// TIA Portal project "Robotic_arm" (V19)

(* hardware
DEVICE "S7-1500/ET200MP station_1"  S7-1500 station
   slot 0: "Rail_0"  Rack  6ES7 590-1***0-0AA0
   slot 1: "PLC_2"  CPU 1511-1 PN  6ES7 511-1AK00-0AB0  V1.8
      slot 3: "CPU display_1"  6ES7591-1AA00-0AA0
      slot 32768: "PROFINET interface_1"  X1
         slot 32769: "Port_1"  X1 P1
         slot 32770: "Port_2"  X1 P2
*)

// ===== PLC "PLC_2"  CPU 1511-1 PN =====

VAR_GLOBAL   // PLC tag table "Cell_IO_list"
   "Cmd_Band_Run" AT %Q0.0 : Bool;
   "Cmd_Gripper_Close" AT %Q0.1 : Bool;
   "Cmd_LoadNew" AT %Q0.2 : Bool;
   "Cmd_Picked" AT %Q0.3 : Bool;
   "Cmd_A1_Pos" AT %QD4 : Real;
   "Cmd_A2_Pos" AT %QD8 : Real;
   "Cmd_A3_Pos" AT %QD12 : Real;
   "Cmd_A4_Pos" AT %QD16 : Real;
   "St_ProductAtPick" AT %I1.0 : Bool;
   "St_Gripper_HasPart" AT %I1.1 : Bool;
   "St_A1_Pos" AT %ID4 : Real;
   "St_A2_Pos" AT %ID8 : Real;
   "St_A3_Pos" AT %ID12 : Real;
   "St_A4_Pos" AT %ID16 : Real;
   "Cmd_Start" AT %M0.0 : Bool;
   "Cmd_Stop" AT %M0.1 : Bool;
   "Cmd_Reset" AT %M0.2 : Bool;
   "Cmd_Auto" AT %M0.3 : Bool;
   "SafeToRun" AT %M0.4 : Bool;
   "Sts_Ready" AT %M10.0 : Bool;
   "Sts_Busy" AT %M10.1 : Bool;
   "Sts_Done" AT %M10.2 : Bool;
   "Sts_Fault" AT %M10.3 : Bool;
   "Sts_State" AT %MW12 : Int;
   "Sts_CycleCount" AT %MW14 : Int;
   "Sts_Hold" AT %M10.4 : Bool;
END_VAR

DATA_BLOCK "DB_RobotPoses"   // DB1
{ S7_Optimized_Access := 'TRUE' }
VERSION : 0.3
   VAR
      HOME_A1 : Real;
      HOME_A2 : Real;
      HOME_A3 : Real;
      HOME_A4 : Real;
      PICK_APP_A1 : Real;
      PICK_APP_A2 : Real := -31.0;
      PICK_APP_A3 : Real := -28.6;
      PICK_APP_A4 : Real := 59.6;
      PICK_A1 : Real;
      PICK_A2 : Real := -50.8;
      PICK_A3 : Real := -24.4;
      PICK_A4 : Real := 75.2;
      PLACE_APP_A1 : Real := 90.0;
      PLACE_APP_A2 : Real := -5.4;
      PLACE_APP_A3 : Real := -51.3;
      PLACE_APP_A4 : Real := 56.7;
      PLACE_A1 : Real := 90.0;
      PLACE_A2 : Real := -42.1;
      PLACE_A3 : Real := -48.1;
      PLACE_A4 : Real := 90.2;
   END_VAR
BEGIN
END_DATA_BLOCK

DATA_BLOCK "iCell"   // DB6
{ S7_Optimized_Access := 'TRUE' }
VERSION : 0.3
// stored: InstanceOfName FB_CellController
"FB_CellController"
BEGIN
END_DATA_BLOCK

FUNCTION_BLOCK "FB_RobotMove"   // FB1, SCL
{ S7_Optimized_Access := 'TRUE' }
VERSION : 0.5
// ----------------------------------------------------------------------------
//  FB_RobotMove : command one joint pose, report Done from NX actual positions
//    - writes the 4 joint set-points to NX (Cmd*)
//    - Done when every joint is within Tol of its target AND a minimum settle
//      time has elapsed.
// 
//    FIX 1: the move re-arms on a rising edge of Execute OR whenever the caller's
//    Step number changes.  The caller passes its own CASE state as Step, so every
//    state transition starts a genuinely new move even when Execute stays TRUE and
//    even when two consecutive states share the same target pose.
//  ----------------------------------------------------------------------------
   VAR_INPUT
      Execute : Bool;
      "Step" : Int;   // caller's state number (FIX 1)
      T1 : Real;   // target joint angles
      T2 : Real;
      T3 : Real;
      T4 : Real;
      Act1 : Real;   // actual angles from NX
      Act2 : Real;
      Act3 : Real;
      Act4 : Real;
      Tol : Real;   // tolerance [deg]
   END_VAR
   VAR_OUTPUT
      Cmd1 : Real := 0.0;   // set-points to NX
      Cmd2 : Real := 0.0;
      Cmd3 : Real := 0.0;
      Cmd4 : Real := 0.0;
      Done : Bool := FALSE;
      Busy : Bool := FALSE;
   END_VAR
   VAR
      prevExec : Bool;
      iBusy : Bool := FALSE;   // FIX 9: internal, so no output is read
      prevStep : Int := -1;
      SettleT : TON_TIME;
   END_VAR
   VAR_TEMP
      inpos : Bool;
      startMove : Bool;
   END_VAR
BEGIN

   // ---- start a new move: rising Execute, or the caller moved to a new step ----
   #startMove := #Execute AND ((NOT #prevExec) OR (#Step <> #prevStep));       // FIX 1

   IF #startMove THEN
       #iBusy := TRUE;
       #Done := FALSE;
   END_IF;

   #prevExec := #Execute;
   #prevStep := #Step;

   // drive set-points only while this move is selected
   IF #Execute THEN
       #Cmd1 := #T1;
       #Cmd2 := #T2;
       #Cmd3 := #T3;
       #Cmd4 := #T4;
   END_IF;

   // in-position test on the NX feedback
   #inpos := (ABS(#Act1 - #T1) <= #Tol) AND
   (ABS(#Act2 - #T2) <= #Tol) AND
   (ABS(#Act3 - #T3) <= #Tol) AND
   (ABS(#Act4 - #T4) <= #Tol);

   // minimum settle / move time.
   // FIX 2: held at IN := FALSE for the re-arm scan, which resets the TON, so the
   //        settle time is honoured for EVERY move and not just the first one.
   #SettleT(IN := #iBusy AND NOT #startMove,
            PT := T#200ms);

   IF #iBusy AND #inpos AND #SettleT.Q THEN
       #Done := TRUE;
       #iBusy := FALSE;
   END_IF;

   // deselecting the move clears it
   IF NOT #Execute THEN
       #Done := FALSE;
       #iBusy := FALSE;
       #prevStep := -1;
   END_IF;

   #Busy := #iBusy;
END_FUNCTION_BLOCK

FUNCTION_BLOCK "FB_Geven"   // FB2, SCL
{ S7_Optimized_Access := 'TRUE' }
VERSION : 0.5
// ----------------------------------------------------------------------------
//  FB_Geven  (GIVE) : run the conveyor until the product reaches the pick
//                     light barrier, then stop the belt. Fault on arrival
//                     time-out (product never arrives).
//    INTERLOCK: the belt only ever runs from inside this module.
//  ----------------------------------------------------------------------------
   VAR_INPUT
      Run : Bool;   // enabled by CellController (active AND not held)
      SafeToRun : Bool;
      St_ProductAtPick : Bool;
   END_VAR
   VAR_OUTPUT
      Cmd_Band_Run : Bool := FALSE;
      Done : Bool := FALSE;
      Fault : Bool := FALSE;
   END_VAR
   VAR
      ArriveTO : TON_TIME;
      iFault : Bool := FALSE;   // FIX 9
      iBand : Bool := FALSE;   // FIX 9
      Cleared : Bool := FALSE;   // FIX 10: barrier seen clear since this module started
   END_VAR
BEGIN

   IF #Run AND #SafeToRun AND NOT #iFault THEN
       IF NOT #Cleared THEN
           // FIX 10: on entry the light barrier may STILL be showing the previous
           //         product (the status signal is one communication step old).
           //         Feed, but do not accept an arrival until the barrier has been
           //         seen clear at least once, so a stale TRUE cannot be mistaken
           //         for the next product arriving.
           #iBand := TRUE;
           #Done := FALSE;
           IF NOT #St_ProductAtPick THEN
               #Cleared := TRUE;
           END_IF;
       ELSIF #St_ProductAtPick THEN
           #iBand := FALSE;     // product detected -> stop belt (pick interlock)
           #Done := TRUE;
       ELSE
           #iBand := TRUE;      // keep feeding
           #Done := FALSE;
       END_IF;
   ELSE
       #iBand := FALSE;
   END_IF;

   // arrival time-out -> representative process error.
   // Called every scan; IN follows the belt command, so it resets by itself when
   // the belt stops or when the module is deselected.
   #ArriveTO(IN := #iBand,
             PT := T#15s);
   IF #ArriveTO.Q THEN
       #iFault := TRUE;
       #iBand := FALSE;
   END_IF;

   IF NOT #Run THEN                  // reset when CellController deselects the module
       #Done := FALSE;
       #iFault := FALSE;
       #Cleared := FALSE;             // FIX 10: re-arm for the next cycle
   END_IF;

   #Cmd_Band_Run := #iBand;
   #Fault := #iFault;
END_FUNCTION_BLOCK

FUNCTION_BLOCK "FB_Verwerken"   // FB3, SCL
{ S7_Optimized_Access := 'TRUE' }
VERSION : 0.3
// RobotCell v0.3 PATCH - only the two blocks that change (FIX 6).
//  FB_RobotMove, FB_Geven, FB_Wegzetten and DB_RobotPoses stay as they are in TIA.
//  ----------------------------------------------------------------------------
//  FB_Verwerken  (PROCESS) : robot picks the product.
//    PICK_APP -> PICK -> close gripper (wait HasPart + 0.5 s) -> lift to PICK_APP
//    -> check the presence sensor is clear (FIX 6).  Missed pick -> retry (max 2).
//    Fault on grip time-out (no part after closing) or on the third missed pick.
//  ----------------------------------------------------------------------------
   VAR_INPUT
      Run : Bool;
      SafeToRun : Bool;
      Act1 : Real;
      Act2 : Real;
      Act3 : Real;
      Act4 : Real;
      St_Gripper_HasPart : Bool;
      St_ProductAtPick : Bool;   // FIX 6: presence sensor at the pick point
   END_VAR
   VAR_OUTPUT
      Cmd1 : Real;
      Cmd2 : Real;
      Cmd3 : Real;
      Cmd4 : Real;
      Cmd_Gripper_Close : Bool;
      Done : Bool;
      Fault : Bool;
      Retries : Int;   // FIX 6: missed picks in this cycle
   END_VAR
   VAR
      State : Int := 0;
      Move : "FB_RobotMove";
      GripTO : TON_TIME;
      GripSettle : TON_TIME;   // FIX 6: jaws settle before lifting
      CheckT : TON_TIME;   // FIX 6: sensor settle after the lift
   END_VAR
BEGIN
   // =====================================================================
   // FB_Verwerken  v0.3  -  CODE ONLY (paste into the code area, replace all)
   //
   // Before pasting, add these 4 lines to the INTERFACE table at the top:
   //   Input   St_ProductAtPick   Bool
   //   Output  Retries            Int
   //   Static  GripSettle         TON_TIME
   //   Static  CheckT             TON_TIME
   // (Run, SafeToRun, Act1..Act4, St_Gripper_HasPart, Cmd1..Cmd4,
   //  Cmd_Gripper_Close, Done, Fault, State, Move, GripTO stay as they are.)
   // =====================================================================

   // FIX 3: the grip time-out is called ONCE PER SCAN, outside the CASE, with an
   //        explicit enable.  It therefore sees IN = FALSE whenever the module is
   //        idle or in another step, which resets it between cycles.  In v0.1 it
   //        was only called from inside CASE 20 with IN := TRUE and kept its
   //        elapsed time, so cycle 2 faulted immediately on entry.
   #GripTO(IN := #Run AND #SafeToRun AND NOT #Fault AND (#State = 20),
           PT := T#3s);
   #GripSettle(IN := #Run AND #SafeToRun AND (#State = 20) AND #St_Gripper_HasPart,
               PT := T#500ms);
   #CheckT(IN := #Run AND #SafeToRun AND (#State = 40),
           PT := T#300ms);

   IF NOT #Run THEN
       #State := 0;
       #Done := FALSE;
       #Fault := FALSE;
       #Retries := 0;
       #Cmd_Gripper_Close := FALSE;
       #Move(Execute := FALSE,
             Step := -1,
             Tol := 1.0,
             Act1 := #Act1,
             Act2 := #Act2,
             Act3 := #Act3,
             Act4 := #Act4);
   ELSIF #SafeToRun AND NOT #Fault THEN
       CASE #State OF
           0:  // move to PICK approach
               #Move(Execute := TRUE,
                     Step := 0,
                     Tol := 1.0,
                     T1 := "DB_RobotPoses".PICK_APP_A1,
                     T2 := "DB_RobotPoses".PICK_APP_A2,
                     T3 := "DB_RobotPoses".PICK_APP_A3,
                     T4 := "DB_RobotPoses".PICK_APP_A4,
                     Act1 := #Act1,
                     Act2 := #Act2,
                     Act3 := #Act3,
                     Act4 := #Act4);
               IF #Move.Done THEN
                   #State := 10;
               END_IF;

           10: // descend to PICK
               #Move(Execute := TRUE,
                     Step := 10,
                     Tol := 1.0,
                     T1 := "DB_RobotPoses".PICK_A1,
                     T2 := "DB_RobotPoses".PICK_A2,
                     T3 := "DB_RobotPoses".PICK_A3,
                     T4 := "DB_RobotPoses".PICK_A4,
                     Act1 := #Act1,
                     Act2 := #Act2,
                     Act3 := #Act3,
                     Act4 := #Act4);
               IF #Move.Done THEN
                   #State := 20;
               END_IF;

           20: // close gripper, wait for part, let the jaws settle (FIX 6)
               #Cmd_Gripper_Close := TRUE;
               IF #GripSettle.Q THEN
                   #State := 30;
               ELSIF #GripTO.Q THEN
                   #Fault := TRUE;            // grip time-out -> error
               END_IF;

           30: // lift back to PICK approach (with part)
               #Move(Execute := TRUE,
                     Step := 30,
                     Tol := 1.0,
                     T1 := "DB_RobotPoses".PICK_APP_A1,
                     T2 := "DB_RobotPoses".PICK_APP_A2,
                     T3 := "DB_RobotPoses".PICK_APP_A3,
                     T4 := "DB_RobotPoses".PICK_APP_A4,
                     Act1 := #Act1,
                     Act2 := #Act2,
                     Act3 := #Act3,
                     Act4 := #Act4);
               IF #Move.Done THEN
                   #State := 40;
               END_IF;

           40: // FIX 6: verify the pick with the presence sensor
               IF #CheckT.Q THEN
                   IF NOT #St_ProductAtPick THEN
                       #State := 100;          // block left the belt -> picked
                   ELSIF #Retries < 2 THEN
                       #Retries := #Retries + 1; // block still there -> missed pick
                       #Cmd_Gripper_Close := FALSE;
                       #State := 50;
                   ELSE
                       #Fault := TRUE;         // third miss -> process error
                   END_IF;
               END_IF;

           50: // FIX 6: retry - open above the block, then descend again
               #Cmd_Gripper_Close := FALSE;
               IF NOT #St_Gripper_HasPart THEN
                   #State := 10;
               END_IF;

           100: // done
               #Done := TRUE;
       END_CASE;
   END_IF;

   // hand the move set-points to the block outputs (read by FB_CellController in step 20)
   #Cmd1 := #Move.Cmd1;
   #Cmd2 := #Move.Cmd2;
   #Cmd3 := #Move.Cmd3;
   #Cmd4 := #Move.Cmd4;
END_FUNCTION_BLOCK

FUNCTION_BLOCK "FB_Wegzetten"   // FB4, SCL
{ S7_Optimized_Access := 'TRUE' }
VERSION : 0.5
// ----------------------------------------------------------------------------
//  FB_Wegzetten  (PUT AWAY) : robot places the product in the storage tray.
//    PLACE_APP -> PLACE -> open gripper (INTERLOCK: only here) -> retract -> HOME.
//  ----------------------------------------------------------------------------
   VAR_INPUT
      Run : Bool;
      SafeToRun : Bool;
      Act1 : Real;
      Act2 : Real;
      Act3 : Real;
      Act4 : Real;
   END_VAR
   VAR_OUTPUT
      Cmd1 : Real := 0.0;
      Cmd2 : Real := 0.0;
      Cmd3 : Real := 0.0;
      Cmd4 : Real := 0.0;
      Cmd_Gripper_Close : Bool := FALSE;
      Done : Bool := FALSE;
      Fault : Bool := FALSE;
   END_VAR
   VAR
      State : Int := 0;
      Mover : "FB_RobotMove";
      OpenT : TON_TIME;
      iFault : Bool := FALSE;   // FIX 9
   END_VAR
BEGIN

   // FIX 3 (same reasoning as FB_Verwerken): called every scan with an explicit
   //        enable so the dwell timer resets between cycles.
   #OpenT(IN := #Run AND #SafeToRun AND NOT #iFault AND (#State = 20),
          PT := T#500ms);

   IF NOT #Run THEN
       #State := 0;
       #Done := FALSE;
       #iFault := FALSE;
       #Cmd_Gripper_Close := TRUE;     // keep holding the part until put-away starts
       #Mover(Execute := FALSE,
              Step := -1,
              Tol := 1.0,
              Act1 := #Act1,
              Act2 := #Act2,
              Act3 := #Act3,
              Act4 := #Act4);
   ELSIF #SafeToRun AND NOT #iFault THEN
       CASE #State OF
           0:  // move to PLACE approach (still holding the part)
               #Cmd_Gripper_Close := TRUE;
               #Mover(Execute := TRUE,
                      Step := 0,
                      Tol := 1.0,
                      T1 := "DB_RobotPoses".PLACE_APP_A1,
                      T2 := "DB_RobotPoses".PLACE_APP_A2,
                      T3 := "DB_RobotPoses".PLACE_APP_A3,
                      T4 := "DB_RobotPoses".PLACE_APP_A4,
                      Act1 := #Act1,
                      Act2 := #Act2,
                      Act3 := #Act3,
                      Act4 := #Act4);
               IF #Mover.Done THEN
                   #State := 10;
               END_IF;

           10: // descend to PLACE
               #Cmd_Gripper_Close := TRUE;
               #Mover(Execute := TRUE,
                      Step := 10,
                      Tol := 1.0,
                      T1 := "DB_RobotPoses".PLACE_A1,
                      T2 := "DB_RobotPoses".PLACE_A2,
                      T3 := "DB_RobotPoses".PLACE_A3,
                      T4 := "DB_RobotPoses".PLACE_A4,
                      Act1 := #Act1,
                      Act2 := #Act2,
                      Act3 := #Act3,
                      Act4 := #Act4);
               IF #Mover.Done THEN
                   #State := 20;
               END_IF;

           20: // open gripper (only allowed above the storage station) + dwell
               #Cmd_Gripper_Close := FALSE;
               IF #OpenT.Q THEN
                   #State := 30;
               END_IF;

           30: // retract to PLACE approach
               #Cmd_Gripper_Close := FALSE;
               #Mover(Execute := TRUE,
                      Step := 30,
                      Tol := 1.0,
                      T1 := "DB_RobotPoses".PLACE_APP_A1,
                      T2 := "DB_RobotPoses".PLACE_APP_A2,
                      T3 := "DB_RobotPoses".PLACE_APP_A3,
                      T4 := "DB_RobotPoses".PLACE_APP_A4,
                      Act1 := #Act1,
                      Act2 := #Act2,
                      Act3 := #Act3,
                      Act4 := #Act4);
               IF #Mover.Done THEN
                   #State := 40;
               END_IF;

           40: // return HOME
               #Cmd_Gripper_Close := FALSE;
               #Mover(Execute := TRUE,
                      Step := 40,
                      Tol := 1.0,
                      T1 := "DB_RobotPoses".HOME_A1,
                      T2 := "DB_RobotPoses".HOME_A2,
                      T3 := "DB_RobotPoses".HOME_A3,
                      T4 := "DB_RobotPoses".HOME_A4,
                      Act1 := #Act1,
                      Act2 := #Act2,
                      Act3 := #Act3,
                      Act4 := #Act4);
               IF #Mover.Done THEN
                   #State := 100;
               END_IF;

           100: // done
               #Cmd_Gripper_Close := FALSE;
               #Done := TRUE;
       END_CASE;
   END_IF;

   // FIX 7: publish the active set-point on the module outputs.  In v0.1 and v0.2
   //        Cmd1..Cmd4 were declared but never assigned, so FB_CellController
   //        multiplexed zeros onto the robot during PROCESS and PUT AWAY.  Placed
   //        after the IF so the outputs also hold the last pose while idle.
   #Cmd1 := #Mover.Cmd1;
   #Cmd2 := #Mover.Cmd2;
   #Cmd3 := #Mover.Cmd3;
   #Cmd4 := #Mover.Cmd4;

   #Fault := #iFault;
END_FUNCTION_BLOCK

FUNCTION_BLOCK "FB_CellController"   // FB5, SCL
{ S7_Optimized_Access := 'TRUE' }
VERSION : 0.3
// ----------------------------------------------------------------------------
//  ----------------------------------------------------------------------------
//  FB_CellController : top sequencer. Coordinates GIVE -> PROCESS -> PUT AWAY,
//    runs CyclesToRun consecutive cycles, handles Auto/Hand, Start/Stop(=Hold)/
//    Reset, aggregates faults, and MUXes the shared robot/gripper/belt outputs
//    so only the active module ever drives NX (single-writer rule).
//  ----------------------------------------------------------------------------
   VAR_INPUT
      Cmd_Start : Bool;
      Cmd_Stop : Bool;   // controlled pause (Hold)
      Cmd_Reset : Bool;
      Cmd_Auto : Bool;   // TRUE = Auto mode, FALSE = Hand
      SafeToRun : Bool;
      CyclesToRun : Int := 3;   // >= 3 consecutive cycles (configurable) feedback from NX / FMU
      St_ProductAtPick : Bool;
      St_Gripper_HasPart : Bool;
      St_A1_Pos : Real;   // commands to NX / FMU
      St_A2_Pos : Real;
      St_A3_Pos : Real;
      St_A4_Pos : Real;
   END_VAR
   VAR_OUTPUT
      Cmd_A1_Pos : Real;
      Cmd_A2_Pos : Real;
      Cmd_A3_Pos : Real;
      Cmd_A4_Pos : Real;
      Cmd_Gripper_Close : Bool;
      Cmd_Band_Run : Bool;
      Cmd_LoadNew : Bool;   // stretched pulse -> FMU spawns next product
      Cmd_Picked : Bool;   // -> FMU freezes product once gripped status to HMI
      Sts_Ready : Bool;
      Sts_Busy : Bool;
      Sts_Done : Bool;
      Sts_Fault : Bool;
      Sts_Hold : Bool;
      Sts_State : Int;
      Sts_CycleCount : Int;
   END_VAR
   VAR
      State : Int := 0;
      Hold : Bool;
      prevStop : Bool;
      LoadReq : Bool;   // FIX 4
      LoadPulse : TON_TIME;   // FIX 4
      Geven : "FB_Geven";
      Verwerken : "FB_Verwerken";
      Wegzetten : "FB_Wegzetten";
   END_VAR
   VAR_TEMP
      gAct : Bool;   // give active
      pAct : Bool;   // process active
      wAct : Bool;   // put-away active
   END_VAR
BEGIN
   // =====================================================================
   // FB_CellController  v0.3  -  CODE ONLY (paste into the code area, replace all)
   //
   // No interface changes.  Compared to your current code only two things differ:
   //   - the #Verwerken(...) call also passes St_ProductAtPick
   //   - step 40: #LoadReq := NOT #St_ProductAtPick   (was TRUE)
   // Compile FB_Verwerken FIRST, then this block.
   // =====================================================================

   // ---- Hold (Stop = controlled pause, Start = resume) ----
   IF #Cmd_Stop AND NOT #prevStop THEN
       #Hold := TRUE;
   END_IF;
   #prevStop := #Cmd_Stop;

   // FIX 5: losing the safety enable, or leaving Auto mode, latches HOLD.  The
   //        cell then requires an explicit Start to continue, so motion never
   //        resumes by itself (safety function SF5, no unexpected restart).
   IF (NOT #SafeToRun) OR (NOT #Cmd_Auto) THEN
       #Hold := TRUE;
   END_IF;

   // Start clears Hold (evaluated last so Start always wins on the same scan)
   IF #Cmd_Start AND #SafeToRun AND #Cmd_Auto THEN
       #Hold := FALSE;
   END_IF;

   // ---- which stage is active this scan ----
   #gAct := (#State = 10);
   #pAct := (#State = 20);
   #wAct := (#State = 30);

   // ---- call all three modules every scan (idle ones reset internally) ----
   #Geven(Run := #gAct AND NOT #Hold,
          SafeToRun := #SafeToRun,
          St_ProductAtPick := #St_ProductAtPick);

   #Verwerken(Run := #pAct,
              SafeToRun := #SafeToRun AND NOT #Hold,
              Act1 := #St_A1_Pos,
              Act2 := #St_A2_Pos,
              Act3 := #St_A3_Pos,
              Act4 := #St_A4_Pos,
              St_Gripper_HasPart := #St_Gripper_HasPart,
              St_ProductAtPick := #St_ProductAtPick);

   #Wegzetten(Run := #wAct,
              SafeToRun := #SafeToRun AND NOT #Hold,
              Act1 := #St_A1_Pos,
              Act2 := #St_A2_Pos,
              Act3 := #St_A3_Pos,
              Act4 := #St_A4_Pos);

   // ---- top sequencer ----
   CASE #State OF
       0:  // INIT / IDLE
           #Sts_Ready := TRUE;
           #Sts_Busy := FALSE;
           #Sts_Done := FALSE;
           #Sts_Fault := FALSE;
           #Cmd_Band_Run := FALSE;
           #Cmd_Gripper_Close := FALSE;
           #Cmd_Picked := FALSE;
           #Cmd_A1_Pos := "DB_RobotPoses".HOME_A1;
           #Cmd_A2_Pos := "DB_RobotPoses".HOME_A2;
           #Cmd_A3_Pos := "DB_RobotPoses".HOME_A3;
           #Cmd_A4_Pos := "DB_RobotPoses".HOME_A4;
           #Sts_CycleCount := 0;
           IF #Cmd_Start AND #Cmd_Auto AND #SafeToRun THEN
               #LoadReq := TRUE;              // spawn first product (FIX 4)
               #State := 10;
           END_IF;

       10: // GIVE
           #Sts_Ready := FALSE;
           #Sts_Busy := TRUE;
           #Cmd_Band_Run := #Geven.Cmd_Band_Run;
           IF #Geven.Fault THEN
               #State := 100;
           END_IF;
           IF #Geven.Done THEN
               #State := 20;
           END_IF;

       20: // PROCESS (pick)
           #Cmd_Band_Run := FALSE;
           #Cmd_A1_Pos := #Verwerken.Cmd1;
           #Cmd_A2_Pos := #Verwerken.Cmd2;
           #Cmd_A3_Pos := #Verwerken.Cmd3;
           #Cmd_A4_Pos := #Verwerken.Cmd4;
           #Cmd_Gripper_Close := #Verwerken.Cmd_Gripper_Close;
           IF #St_Gripper_HasPart THEN
               #Cmd_Picked := TRUE;
           END_IF;   // freeze product in FMU
           IF #Verwerken.Fault THEN
               #State := 100;
           END_IF;
           IF #Verwerken.Done THEN
               #State := 30;
           END_IF;

       30: // PUT AWAY (place)
           #Cmd_A1_Pos := #Wegzetten.Cmd1;
           #Cmd_A2_Pos := #Wegzetten.Cmd2;
           #Cmd_A3_Pos := #Wegzetten.Cmd3;
           #Cmd_A4_Pos := #Wegzetten.Cmd4;
           #Cmd_Gripper_Close := #Wegzetten.Cmd_Gripper_Close;
           IF #Wegzetten.Fault THEN
               #State := 100;
           END_IF;
           IF #Wegzetten.Done THEN
               #State := 40;
           END_IF;

       40: // CYCLE END
           #Sts_CycleCount := #Sts_CycleCount + 1;
           #Cmd_Picked := FALSE;
           IF #Sts_CycleCount < #CyclesToRun THEN
               #LoadReq := NOT #St_ProductAtPick;  // FIX 6: next product only if the pick is clear
               #State := 10;
           ELSE
               #State := 50;
           END_IF;

       50: // ALL CYCLES DONE
           #Sts_Busy := FALSE;
           #Sts_Done := TRUE;
           #Cmd_Band_Run := FALSE;
           IF #Cmd_Reset THEN
               #State := 0;
           END_IF;

       100: // FAULT (safe state)
           #Sts_Busy := FALSE;
           #Sts_Fault := TRUE;
           #Cmd_Band_Run := FALSE;           // belt off
           // robot holds last commanded pose; gripper keeps its state
           IF #Cmd_Reset THEN
               #Sts_Fault := FALSE;
               #State := 0;
           END_IF;
   END_CASE;

   // ---- FIX 4: stretch Cmd_LoadNew so the co-simulation cannot miss it ----
   #LoadPulse(IN := #LoadReq,
              PT := T#200ms);
   IF #LoadPulse.Q THEN
       #LoadReq := FALSE;
   END_IF;
   #Cmd_LoadNew := #LoadReq;

   // ---- Hold overlay: freeze robot at current actual + stop belt ----
   IF #Hold AND (#State >= 10) AND (#State <= 30) THEN
       #Cmd_Band_Run := FALSE;
       #Cmd_A1_Pos := #St_A1_Pos;
       #Cmd_A2_Pos := #St_A2_Pos;
       #Cmd_A3_Pos := #St_A3_Pos;
       #Cmd_A4_Pos := #St_A4_Pos;
   END_IF;

   #Sts_Hold := #Hold;
   #Sts_State := #State;
END_FUNCTION_BLOCK

ORGANIZATION_BLOCK "Main"   // OB1, SCL, ProgramCycle
TITLE = "Main Program Sweep (Cycle)"
{ S7_Optimized_Access := 'TRUE' }
VERSION : 0.1
   VAR_INPUT
      Initial_Call : Bool;   // Initial call of this OB
      Remanence : Bool;   // =True, if remanent data are available
   END_VAR
BEGIN
   // ============================================================================
   //  Main [OB1] - top-level call of the pick-&-place cell
   //  Paste the block below into an SCL organization block named "Main".
   //
   //    :=  passes a tag INTO the function block   (inputs)
   //    =>  writes a function block output OUT to a tag
   //
   //  Every line ends with a comma except the last, which closes with  );
   //  All 27 parameters are wired.  Sts_Hold needs the %M10.4 tag in Cell_IO_list.
   // ============================================================================

   "iCell"(Cmd_Start := "Cmd_Start",
           Cmd_Stop := "Cmd_Stop",
           Cmd_Reset := "Cmd_Reset",
           Cmd_Auto := "Cmd_Auto",
           SafeToRun := "SafeToRun",
           CyclesToRun := 3,
           St_ProductAtPick := "St_ProductAtPick",
           St_Gripper_HasPart := "St_Gripper_HasPart",
           St_A1_Pos := "St_A1_Pos",
           St_A2_Pos := "St_A2_Pos",
           St_A3_Pos := "St_A3_Pos",
           St_A4_Pos := "St_A4_Pos",
           Cmd_A1_Pos => "Cmd_A1_Pos",
           Cmd_A2_Pos => "Cmd_A2_Pos",
           Cmd_A3_Pos => "Cmd_A3_Pos",
           Cmd_A4_Pos => "Cmd_A4_Pos",
           Cmd_Gripper_Close => "Cmd_Gripper_Close",
           Cmd_Band_Run => "Cmd_Band_Run",
           Cmd_LoadNew => "Cmd_LoadNew",
           Cmd_Picked => "Cmd_Picked",
           Sts_Ready => "Sts_Ready",
           Sts_Busy => "Sts_Busy",
           Sts_Done => "Sts_Done",
           Sts_Fault => "Sts_Fault",
           Sts_Hold => "Sts_Hold",
           Sts_State => "Sts_State",
           Sts_CycleCount => "Sts_CycleCount");
END_ORGANIZATION_BLOCK